// TIA Portal V21 export
FUNCTION_BLOCK "GraphQualification"   // FB, GRAPH
// stored: AutoNumber true
   VAR_INPUT
      ACK_EF : Bool;
      StartCommand : Bool;
      ResetCommand : Bool;
      GuardClosed : Bool;
      SupervisionTrip : Bool;
   END_VAR
   VAR_OUTPUT
      MotorA : Bool;
      MotorB : Bool;
   END_VAR
BEGIN
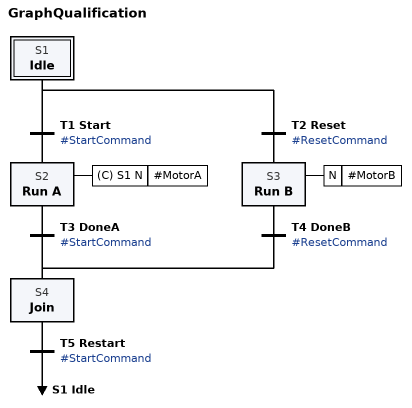
   // sequencer 1: Parallel cycle / Paralleler Ablauf
   INITIAL_STEP Idle:   // S1
      interlock C := #GuardClosed;
      supervision V := #SupervisionTrip;
   END_STEP
   TRANSITION Start FROM Idle TO "Run A"   // T1
      := #StartCommand;
   END_TRANSITION
   TRANSITION Reset FROM Idle TO "Run B"   // T2
      := #ResetCommand;
   END_TRANSITION
   STEP "Run A":   // S2, max time T#10s, warning time T#8s
      interlock C := #GuardClosed;
      supervision V := #SupervisionTrip;   // Travel timeout
      (C) S1  N    #MotorA
   END_STEP
   TRANSITION DoneA FROM "Run A" TO Join   // T3
      := #StartCommand;
   END_TRANSITION
   STEP "Run B":   // S3
      interlock C := #GuardClosed;
      supervision V := #SupervisionTrip;
              N    #MotorB
   END_STEP
   TRANSITION DoneB FROM "Run B" TO Join   // T4
      := #ResetCommand;
   END_TRANSITION
   STEP Join:   // S4
      interlock C := #GuardClosed;
      supervision V := #SupervisionTrip;
   END_STEP
   TRANSITION Restart FROM Join TO Idle   // T5, jump
      := #StartCommand;
   END_TRANSITION
END_FUNCTION_BLOCK
